Fanuc KAREL source: kt00330.KL

-- PROVISIONAL review KL for V1013-1; original PC SHA256 5e981b51c005414e045c2f6e82742cad737363c2fc9916c964a3919b62253e23
-- Incomplete behavior may be omitted. Consult companion uncertainty JSON. Do not deploy.
PROGRAM KT00330
%NOLOCKGROUP
VAR
  I1 : INTEGER
  R2 : REAL
  OUT : BOOLEAN
BEGIN
  -- UNRESOLVED_PC offsets 5-16; opcodes 2E,23
  -- UNRESOLVED_PC offsets 21-32; opcodes 2E,23
  -- UNRESOLVED_PC offsets 37-59; opcodes 21,21,29,64,29,6F,23
  -- UNRESOLVED_PC offsets 64-68; opcodes 7F
END KT00330
